// TIA Portal V20 export
DATA_BLOCK "T12_Resultado"   // DB48901
{ S7_Optimized_Access := 'TRUE' }
AUTHOR : IA
FAMILY : PRUEBA
VERSION : 0.1
// Tanda 7: un Bool por prueba
// stored: AutoNumber false
   VAR
      L_Constante : Bool;   // VAR CONSTANT en un FB KOP (LIMITE = 10)
      L_Variant : Bool;   // Variant como entrada de un FB KOP + VariantGet
      S_ArrayStar : Bool;   // Array[*] en SCL: suma con LOWER_BOUND/UPPER_BOUND de un Array[0..4] y de un Array[1..3]
      L_ArrayStar : Bool;   // Array[*] en la interfaz de una FC KOP (SD) llamada con dos arrays
      L_Startup : Bool;   // OB100 (Startup) creado por XML: se ha ejecutado al arrancar
      L_ProgError : Bool;   // OB121 (ProgrammingError) creado por XML: atrapa un índice fuera de rango
      Vida : DInt;   // Sube cada ciclo
      OK : Int;   // Correctas
      Total : Int := 6;   // Pruebas
      Todo_OK : Bool;   // Todas correctas
   END_VAR
BEGIN
END_DATA_BLOCK
